(* CoDeSys 2.3 export: translation.exp *)

(* POU PLC_LD_PRG_TR, FAI *)
PROGRAM PLC_LD_PRG_TR
VAR
END_VAR
(* body not read: x-want_COMMENT *)
END_PROGRAM
